// TIA Portal V20 export
// export: Created 2026-11-18T05:23:18.8006841Z, ExportSetting WithDefaults, DisplayName Totally Integrated Automation Portal, DisplayVersion V20 Update 7, DisplayName TIA Portal Openness, DisplayVersion V20 Update 7, DisplayName TIA Portal Version Control Interface, DisplayVersion V20 Update 7, DisplayName TIA Portal Test Suite Advanced, DisplayVersion V20, DisplayName SINAMICS Startdrive Advanced, DisplayVersion V20 SP1 Update 1, DisplayName SINAMICS Startdrive G110M, G120, G120C, G120D, G120P, G115D, DisplayVersion V20 SP1 Update 1, DisplayName SINAMICS Startdrive G130, G150, S120, S150, SINAMICS MV, G220, S200, S210, DisplayVersion V20 SP1 Update 1, DisplayName STEP 7 Professional, DisplayVersion V20 Update 7, DisplayName STEP 7 Safety, DisplayVersion V20 Update 2, DisplayName WinCC Basic/Comfort/Advanced, DisplayVersion V20 Update 7, DisplayName WinCC Unified, DisplayVersion V20 Update 7
DATA_BLOCK "zzE2eFbI_DB"   // DB16
VERSION : 0.1
// stored: AutoNumber true, DBAccessibleFromOPCUA true, DBAccessibleFromWebserver true, InstanceOfName zzE2eFbI, InstanceOfType FB
"zzE2eFbI"
   // VAR_INPUT
   //    inV : Int := 5;
   //    inW : Int;
   // END_VAR
   // VAR
   //    stV : Int;
   //    stU { S7_SetPoint := 'True'} : "zzE2eUdtA";
   // END_VAR
BEGIN
   stU.as[*].x := 1;   // as x
END_DATA_BLOCK
